Fanuc KAREL source: kt00712.KL

-- PROVISIONAL review KL for V1013-1; original PC SHA256 45168bbdca7b1484686899e4d8b2fd1577fb150ec00b2e1d599ca7b52dba0e2a
-- Incomplete behavior may be omitted. Consult companion uncertainty JSON. Do not deploy.
PROGRAM KT00712
%NOLOCKGROUP
VAR
  S1 : STRING[80]
  S2 : STRING[80]
  OUT : BOOLEAN
BEGIN
  -- UNRESOLVED_PC offsets 5-14; opcodes 3F,75
  -- UNRESOLVED_PC offsets 19-28; opcodes 3F,75
  -- UNRESOLVED_PC offsets 33-42; opcodes 3F,75
  -- UNRESOLVED_PC offsets 47-56; opcodes 3F,75
  -- UNRESOLVED_PC offsets 61-76; opcodes 22,63,23
  -- UNRESOLVED_PC offsets 81-85; opcodes 7F
END KT00712
